Staubli VAL3: simulate.pjx

--- simulate.pjx ---
Parameters version=s8.10.3Cs9_BS2093 stackSize=5000 millimeterUnit=true
Program file=goHome.pgx
Program file=simulate_UI.pgx
Program file=simulateHome.pgx
Program file=simulatePROG.pgx
Program file=simulateTRAJ.pgx
Program file=start.pgx
Program file=stop.pgx
Data file=simulate.dtx
Library alias=savedata path=Disk://source/saveData/saveData.pjx
Library alias=rs path=Disk://source/projectSource/robotStatus/robotStatus.pjx
Library alias=util path=Disk://HMI_cs9/HMI_util/HMI_util.pjx
Library alias=trajectory path=Disk://source/projectSource/trajectory/trajectory.pjx
Library alias=program path=Disk://source/projectSource/program/program.pjx

--- simulate.dtx ---
mdesc mNomSpeed
mdesc mSimulate = {accel=64, vel=80, decel=64, blend=off}
string sMsg
bool bCancel

--- start.pgx ---
program start()
begin
end

--- goHome.pgx ---
public program goHome()
begin
  //stopMove()
  if !isEmpty()
    resetMotion()
  endIf
  movej(herej(),flange,mSimulate)
  movej(savedata:jHome,flange,mSimulate)
  waitEndMove()
end

--- simulate_UI.pgx ---
program simulate_UI()
  local bool l_bExit
begin

  do
    if util:sPage!="simulate"
      util:sPage="simulate"
      userPageBind("simulate","lbl2","innerHTML",sMsg,1,"r")
      userPageBindClick("simulate","img1",bCancel,true)
      userPage("simulate")
      delay(0.1)
    endIf
    sMsg=rs:sTrajStatus
    if bCancel
      bCancel=false
      l_bExit=true
    endIf


    delay(0)
  until l_bExit==true or taskStatus("simulate")==-1
  rs:bSimulate=false
  rs:bGOTO=false
  if taskStatus("simulate")>-1
    taskKill("simulate")
    resetMotion()
  endIf

end

--- simulateHome.pgx ---
public program simulateHome()
  local bool l_bResult
  local bool l_bExit
begin
  if !rs:bIsCycle and workingMode()==1
    l_bResult=userPageConfirm("是否移动到Home位置？")
    if l_bResult
      rs:bSimulate=true

      taskCreate "simulate",50,goHome()
      sMsg="回Home过程。。。"
      call simulate_UI()
    endIf
  else
    userPageAlert("条件不满足：不再生产周期&切换到手动模式")
  endIf
end

--- simulatePROG.pgx ---
public program simulatePROG(string x_sKey)
  local bool l_bResult
begin
  if !rs:bIsCycle and workingMode()==1
    l_bResult=userPageConfirm("是否模拟PROG："+x_sKey+"？")
    if l_bResult
      resetMotion()
      rs:bGOTO=false
      rs:bSimulate=true
      //添加traj任务‘
      taskCreate "simulate",100,program:makeTraj(x_sKey)
      //
      sMsg="模拟PROG过程。。。"
      sMsg=rs:sTrajStatus
      call simulate_UI()
    endIf
  else
    userPageAlert("条件不满足：不再生产周期&切换到手动模式")
  endIf
end

--- simulateTRAJ.pgx ---
public program simulateTRAJ(string x_sKey)
  local bool l_bResult
begin
  if !rs:bIsCycle and workingMode()==1
    l_bResult=userPageConfirm("是否模拟TRAJ："+x_sKey+"？")
    if l_bResult
      resetMotion()
      rs:bSimulate=true
      rs:bGOTO=false
      //添加traj任务‘
      taskCreate "simulate",100,trajectory:makeTraj(x_sKey)
      //
      sMsg="模拟TRAJ过程。。。"
      sMsg=rs:sTrajStatus
      call simulate_UI()
    endIf
  else
    userPageAlert("条件不满足：不再生产周期&切换到手动模式")
  endIf
end

--- stop.pgx ---
program stop()
begin
end
